Universal Robots URScript: T009_deepseek-coder-v2_16b-lite-instruct-q4_K_M_baseline_rep1.urscript

# Define the home position
def home_position():
    movej([0.0, -1.8, 1.8, -1.5, 1.5, 0.0], 180, 0.01, 0.01)

# Move to the above scan start position
def move_above_scan_start():
    movej([0.0, -1.8, 1.8, -1.5, 1.5, 0.0], 150, 0.01, 0.01)

# Move to the descend to scan height position
def move_descend_to_scan_height():
    movej([0.0, -1.8, 1.8, -1.5, 1.5, 0.0], 80, 0.01, 0.01)

# Move to the scan line 1 position
def move_scan_line_1():
    movej([0.0, -1.8, 1.8, -1.5, 1.5, 0.0], 50, 0.01, 0.01)

# Move to the step to line 2 position
def move_step_to_line_2():
    movej([0.0, -1.8, 1.8, -1.5, 1.5, 0.0], 80, 0.01, 0.01)

# Define the sequence of moves
def laser_surface_scan():
    home_position()
    move_above_scan_start()
    move_descend_to_scan_height()
    move_scan_line_1()
    move_step_to_line_2()
    # Continue with the rest of the sequence...

# Call the laser surface scan function
laser_surface_scan()
